// TIA Portal V19 export
// export: Created 2026-10-15T10:10:37.454039Z, ExportSetting WithDefaults, DisplayName Totally Integrated Automation Portal, DisplayVersion V19, DisplayName TIA Portal Openness, DisplayVersion V19, DisplayName TIA Portal Version Control Interface, DisplayVersion V19, DisplayName STEP 7 Professional, DisplayVersion V19, DisplayName STEP 7 Safety, DisplayVersion V19, DisplayName WinCC Basic/Comfort/Advanced, DisplayVersion V19, DisplayName WinCC Unified, DisplayVersion V19
ORGANIZATION_BLOCK "OB100"   // OB100, SCL, Startup
TITLE = "Complete Restart"
{ S7_Optimized_Access := 'TRUE' }
VERSION : 0.1
// stored: AutoNumber true, IsIECCheckEnabled false, SetENOAutomatically false
   VAR_INPUT
      LostRetentive : Bool;   // True if retentive data are lost
      LostRTC : Bool;   // True if date and time are lost
   END_VAR
   VAR_TEMP
      n : Int;
   END_VAR
BEGIN

   // RE plus RS120 bit 3: all M retained. Default T/Z 0..63 retained.
   FOR #n := 64 TO 127 DO
       "ROLL_State".S5Timers[#n].RemainingMs := 0.0;
       "ROLL_State".S5Timers[#n].BaseMs := 0;
       "ROLL_State".S5Timers[#n].Mode := 0;
       "ROLL_State".S5Timers[#n].Q := FALSE;
       "ROLL_State".S5Timers[#n].Previous := FALSE;
       "ROLL_State".S5Counters[#n].Value := 0;
       "ROLL_State".S5Counters[#n].SetPrevious := FALSE;
       "ROLL_State".S5Counters[#n].UpPrevious := FALSE;
       "ROLL_State".S5Counters[#n].DownPrevious := FALSE;
   END_FOR;
   "ROLL_IO".FirstCycle := TRUE;
   "ROLL_IO".ClockMs := 0.0;
   "ROLL_IO".RuntimeMemory := 0.0;
   "ROLL_IO".PhysicalOutputsEnabled := FALSE;
   "ROLL_HMI".Connected := FALSE;
   "ROLL_State".M[0, 1] := TRUE;
   "ROLL_State".M[0, 2] := TRUE;
   "ROLL_State".M[191, 0] := TRUE;
   "ROLL_State".M[190, 5] := FALSE;
   "ROLL_State".M[190, 6] := FALSE;
   "ROLL_State".M[190, 1] := TRUE;
   "ROLL_State".M[191, 4] := TRUE;
   "ROLL_FB90"();
   "ROLL_ShowRecipe"();
END_ORGANIZATION_BLOCK
